(* PLC project probe.project, CODESYS CODESYS V3.5 SP17 Patch 3 *)
(* stored: creationDateTime 2026-10-20T03:54:26.7441148, modificationDateTime 1601-01-01T03:00:00 *)

FUNCTION_BLOCK FB_ProbeSt
  VAR_INPUT
    xIn : BOOL;
  END_VAR
  VAR_OUTPUT
    xQ : BOOL;
    iCount : INT;
  END_VAR
  VAR
    fbTon : TON;
    fbEdge : R_TRIG;
  END_VAR

            fbTon(IN := xIn, PT := T#1S);
xQ := fbTon.Q;
fbEdge(CLK := xIn);
IF fbEdge.Q THEN
    iCount := iCount + 1;
END_IF

          
END_FUNCTION_BLOCK
